(* PLC project Storage_Main, Beckhoff Automation GmbH TwinCAT PLC Control 3.5.13.21 *)
(* stored: creationDateTime 2026-11-24T10:30:00, modificationDateTime 2026-11-24T10:30:00 *)

PROGRAM SFC_Sequence
// =====================================================================
// SFC_Sequence (Sequential Function Chart)
// Homing and the automatic sequence (GRAFCET E70 .. S70).
// Called from MAIN every cycle. All variables are in MAIN (MAIN.xxx).
// Every step has one ST action (<step>_Active) that runs while the step is active.
// The motors are switched off in MAIN before this chart is called, so a step
// only has to switch ON what it needs.
// =====================================================================
VAR_INPUT
    SFCReset : BOOL;            // SFC flag: TRUE = chart back to the initial step S0 (STOP / homing timeout)
END_VAR
VAR
END_VAR

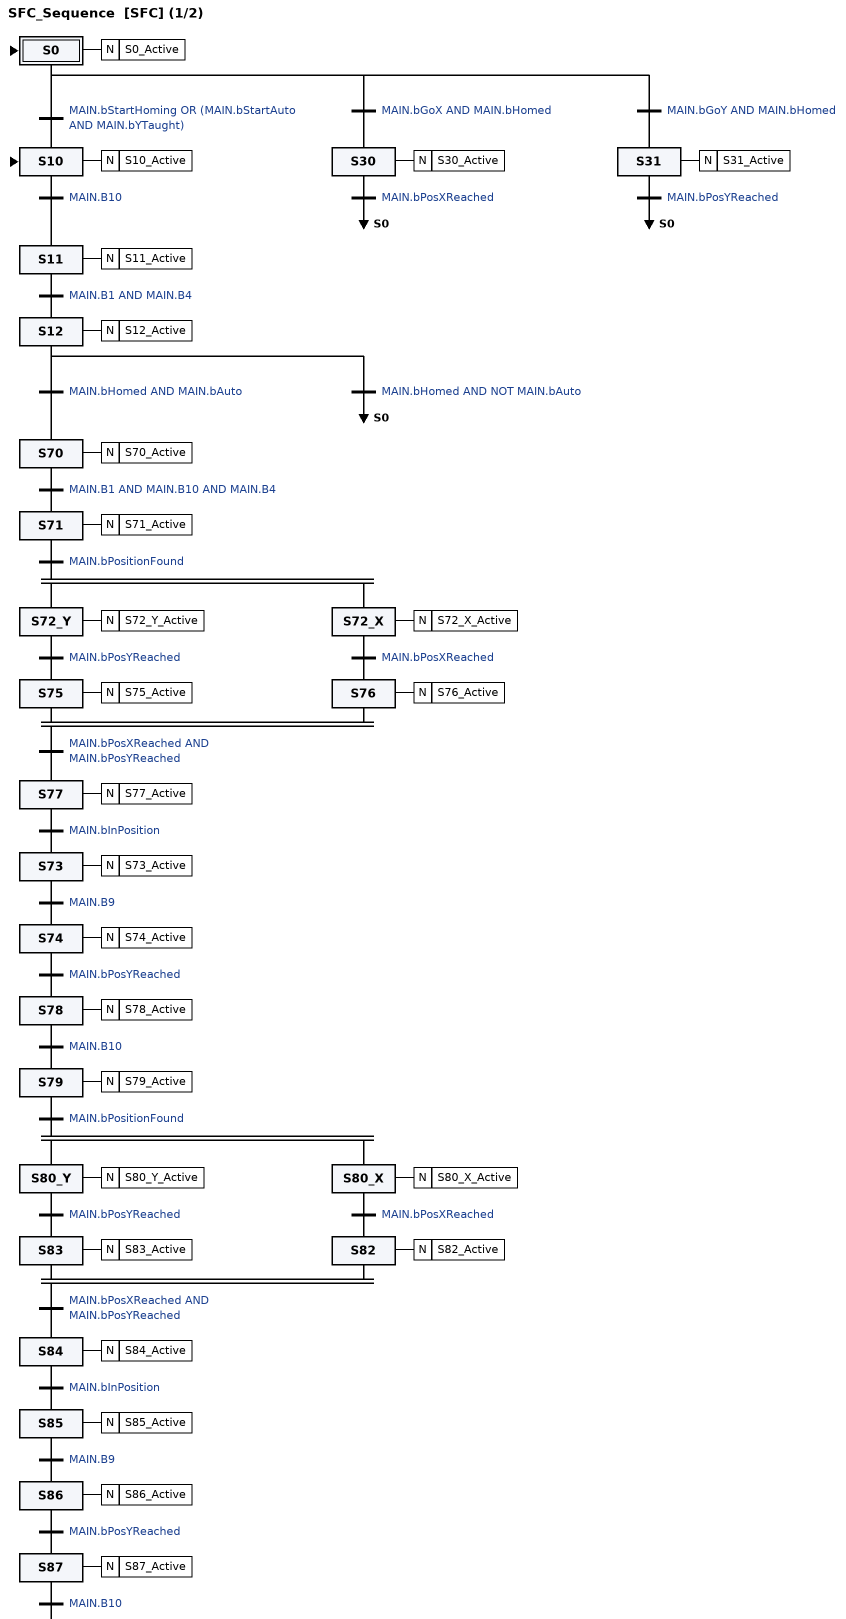
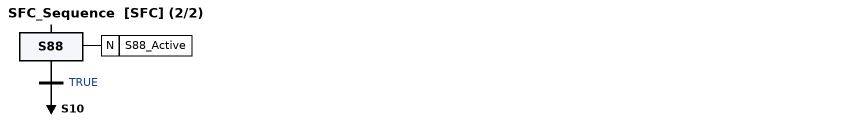
INITIAL_STEP S0:
  S0_Active(N);
END_STEP
TRANSITION FROM S0 TO S10
  := MAIN.bStartHoming OR (MAIN.bStartAuto AND MAIN.bYTaught);
END_TRANSITION
TRANSITION FROM S0 TO S30
  := MAIN.bGoX AND MAIN.bHomed;
END_TRANSITION
TRANSITION FROM S0 TO S31
  := MAIN.bGoY AND MAIN.bHomed;
END_TRANSITION
STEP S10:
  S10_Active(N);
END_STEP
TRANSITION FROM S10 TO S11
  := MAIN.B10;
END_TRANSITION
STEP S11:
  S11_Active(N);
END_STEP
TRANSITION FROM S11 TO S12
  := MAIN.B1 AND MAIN.B4;
END_TRANSITION
STEP S12:
  S12_Active(N);
END_STEP
TRANSITION FROM S12 TO S70
  := MAIN.bHomed AND MAIN.bAuto;
END_TRANSITION
TRANSITION FROM S12 TO S0
  := MAIN.bHomed AND NOT MAIN.bAuto;
END_TRANSITION
STEP S70:
  S70_Active(N);
END_STEP
TRANSITION FROM S70 TO S71
  := MAIN.B1 AND MAIN.B10 AND MAIN.B4;
END_TRANSITION
STEP S71:
  S71_Active(N);
END_STEP
TRANSITION FROM S71 TO (S72_Y, S72_X)
  := MAIN.bPositionFound;
END_TRANSITION
STEP S72_Y:
  S72_Y_Active(N);
END_STEP
TRANSITION FROM S72_Y TO S75
  := MAIN.bPosYReached;
END_TRANSITION
STEP S75:
  S75_Active(N);
END_STEP
TRANSITION FROM (S75, S76) TO S77
  := MAIN.bPosXReached AND MAIN.bPosYReached;
END_TRANSITION
STEP S72_X:
  S72_X_Active(N);
END_STEP
TRANSITION FROM S72_X TO S76
  := MAIN.bPosXReached;
END_TRANSITION
STEP S76:
  S76_Active(N);
END_STEP
STEP S77:
  S77_Active(N);
END_STEP
TRANSITION FROM S77 TO S73
  := MAIN.bInPosition;
END_TRANSITION
STEP S73:
  S73_Active(N);
END_STEP
TRANSITION FROM S73 TO S74
  := MAIN.B9;
END_TRANSITION
STEP S74:
  S74_Active(N);
END_STEP
TRANSITION FROM S74 TO S78
  := MAIN.bPosYReached;
END_TRANSITION
STEP S78:
  S78_Active(N);
END_STEP
TRANSITION FROM S78 TO S79
  := MAIN.B10;
END_TRANSITION
STEP S79:
  S79_Active(N);
END_STEP
TRANSITION FROM S79 TO (S80_Y, S80_X)
  := MAIN.bPositionFound;
END_TRANSITION
STEP S80_Y:
  S80_Y_Active(N);
END_STEP
TRANSITION FROM S80_Y TO S83
  := MAIN.bPosYReached;
END_TRANSITION
STEP S83:
  S83_Active(N);
END_STEP
TRANSITION FROM (S83, S82) TO S84
  := MAIN.bPosXReached AND MAIN.bPosYReached;
END_TRANSITION
STEP S80_X:
  S80_X_Active(N);
END_STEP
TRANSITION FROM S80_X TO S82
  := MAIN.bPosXReached;
END_TRANSITION
STEP S82:
  S82_Active(N);
END_STEP
STEP S84:
  S84_Active(N);
END_STEP
TRANSITION FROM S84 TO S85
  := MAIN.bInPosition;
END_TRANSITION
STEP S85:
  S85_Active(N);
END_STEP
TRANSITION FROM S85 TO S86
  := MAIN.B9;
END_TRANSITION
STEP S86:
  S86_Active(N);
END_STEP
TRANSITION FROM S86 TO S87
  := MAIN.bPosYReached;
END_TRANSITION
STEP S87:
  S87_Active(N);
END_STEP
TRANSITION FROM S87 TO S88
  := MAIN.B10;
END_TRANSITION
STEP S88:
  S88_Active(N);
END_STEP
TRANSITION FROM S88 TO S10
  := TRUE;
END_TRANSITION
STEP S30:
  S30_Active(N);
END_STEP
TRANSITION FROM S30 TO S0
  := MAIN.bPosXReached;
END_TRANSITION
STEP S31:
  S31_Active(N);
END_STEP
TRANSITION FROM S31 TO S0
  := MAIN.bPosYReached;
END_TRANSITION

ACTION S0_Active:
                // S0: Manual mode (initial step)
// Jog, teach and the commands are handled in MAIN (ST) while nStep = 0.
MAIN.nStep := 0;
              
END_ACTION

ACTION S10_Active:
                // S10: Homing - arm back (until B10)
MAIN.nStep := 10;
MAIN.bHomed := FALSE;
MAIN.M4_Back := TRUE;
              
END_ACTION

ACTION S11_Active:
                // S11: Homing - X to B1 and Y to B4 at the same time
MAIN.nStep := 11;
MAIN.M2_Back := NOT MAIN.B1;                     // each axis stops at its own switch
MAIN.M3_Up   := NOT MAIN.B4;
              
END_ACTION

ACTION S12_Active:
                // S12: Homing - wait 0.5 s (tonSettle in MAIN), then set both positions to 0
MAIN.nStep := 12;
IF MAIN.tonSettle.Q THEN
    MAIN.nPosX := 0;
    MAIN.nPosY := 0;
    MAIN.bHomed := TRUE;
END_IF
              
END_ACTION

ACTION S70_Active:
                // S70 = E70 Entry step: wait until the crane is at home (B1 * B10 * B4)
MAIN.nStep := 70;
MAIN.bShelfSelected := FALSE;                    // ignore any old shelf selection
              
END_ACTION

ACTION S71_Active:
                // S71: Get PosX and PosY from the arrays according to the operator's choice
// (nStep = 71 shows the 3x3 shelf selection on the HMI)
MAIN.nStep := 71;
MAIN.bPosXReached := FALSE;
MAIN.bPosYReached := FALSE;

IF MAIN.bShelfSelected THEN
    MAIN.bShelfSelected := FALSE;
    IF MAIN.nSelColumn >= 1 AND MAIN.nSelColumn <= 3 AND MAIN.nSelRow >= 1 AND MAIN.nSelRow <= 3 THEN
        MAIN.nTargetX := MAIN.xPosition[MAIN.nSelColumn];
        MAIN.nTargetY := MAIN.yPosition[MAIN.nSelRow];
        MAIN.bPositionFound := TRUE;
    END_IF
END_IF
              
END_ACTION

ACTION S72_Y_Active:
                // S72 (Y part): Y moves to the shelf height (M3_Down via ACT_Positioning)
MAIN.nStep := 72;
MAIN.bPositionFound := FALSE;
MAIN.bDriveY := TRUE;
              
END_ACTION

ACTION S75_Active:
                // S75: Y in position (M3 off), waits for X
MAIN.nStep := 75;
              
END_ACTION

ACTION S72_X_Active:
                // S72 (X part): X moves to the shelf column (M2_Forward via ACT_Positioning)
MAIN.nStep := 72;
MAIN.bPositionFound := FALSE;
MAIN.bDriveX := TRUE;
              
END_ACTION

ACTION S76_Active:
                // S76: X in position (M2 off), waits for Y
MAIN.nStep := 76;
              
END_ACTION

ACTION S77_Active:
                // S77: Both axes in position
MAIN.nStep := 77;
MAIN.bInPosition := TRUE;
              
END_ACTION

ACTION S73_Active:
                // S73: Arm out under the pallet (until B9)
MAIN.nStep := 73;
MAIN.M4_Forward := TRUE;
MAIN.bInPosition := FALSE;
MAIN.nTargetY := MAIN.yPosition[MAIN.nSelRow] - MAIN.nLiftOffset;   // prepare the lift (up = smaller Y)
MAIN.bPosYReached := FALSE;
              
END_ACTION

ACTION S74_Active:
                // S74: Lift the pallet off the shelf (M3_Up via ACT_Positioning)
MAIN.nStep := 74;
MAIN.bDriveY := TRUE;
              
END_ACTION

ACTION S78_Active:
                // S78: Arm back with the pallet (until B10)
MAIN.nStep := 78;
MAIN.M4_Back := TRUE;
              
END_ACTION

ACTION S79_Active:
                // S79: Get the delivery position (index 0 = conveyor)
MAIN.nStep := 79;
MAIN.nTargetX := MAIN.xPosition[0];              // DeliveryPosX
MAIN.nTargetY := MAIN.yPosition[0];              // DeliveryPosY
MAIN.bPosXReached := FALSE;
MAIN.bPosYReached := FALSE;
MAIN.bPositionFound := TRUE;
              
END_ACTION

ACTION S80_Y_Active:
                // S80/S81 (Y part): Y moves up or down to the delivery height.
// ACT_Positioning chooses the direction (M3_Up or M3_Down) by itself.
MAIN.nStep := 80;
MAIN.bPositionFound := FALSE;
MAIN.bDriveY := TRUE;
              
END_ACTION

ACTION S83_Active:
                // S83: Y in position (M3 off), waits for X
MAIN.nStep := 83;
              
END_ACTION

ACTION S80_X_Active:
                // S80/S81 (X part): X moves back to the conveyor (M2_Back via ACT_Positioning)
MAIN.nStep := 80;
MAIN.bPositionFound := FALSE;
MAIN.bDriveX := TRUE;
              
END_ACTION

ACTION S82_Active:
                // S82: X in position (M2 off), waits for Y
MAIN.nStep := 82;
              
END_ACTION

ACTION S84_Active:
                // S84: Both axes in position
MAIN.nStep := 84;
MAIN.bInPosition := TRUE;
              
END_ACTION

ACTION S85_Active:
                // S85: Arm out over the conveyor (until B9)
MAIN.nStep := 85;
MAIN.M4_Forward := TRUE;
MAIN.bInPosition := FALSE;
MAIN.nTargetY := MAIN.yPosition[0] + MAIN.nLowerOffset;   // prepare lowering (down = larger Y)
MAIN.bPosYReached := FALSE;
              
END_ACTION

ACTION S86_Active:
                // S86: Lower the pallet onto the conveyor (M3_Down via ACT_Positioning)
MAIN.nStep := 86;
MAIN.bDriveY := TRUE;
              
END_ACTION

ACTION S87_Active:
                // S87: Arm back (until B10)
MAIN.nStep := 87;
MAIN.M4_Back := TRUE;
              
END_ACTION

ACTION S88_Active:
                // S88 = S70 Exit step: home again. Homing returns to S70 because bAuto is still TRUE.
MAIN.nStep := 88;
              
END_ACTION

ACTION S30_Active:
                // S30: Manual - move X to xPosition[nTeachSlot] (target set in ACT_Manual)
MAIN.nStep := 30;
MAIN.bDriveX := TRUE;
              
END_ACTION

ACTION S31_Active:
                // S31: Manual - move Y to yPosition[nTeachSlot] (target set in ACT_Manual)
MAIN.nStep := 31;
MAIN.bDriveY := TRUE;
              
END_ACTION
END_PROGRAM
